SUBAPPLICATION logiBUS_QXA_OPC (* logiBUS DQ Kanal: OPC-UA Read/Write (generisch, ein Kanal, ohne VT-Button/Hintergrundfarbe - fuer Module ohne ISOBUS/VT-Anbindung) *)
  (* Standard: 61499-2 *)
  (* Version 1.0, 2026-08-27, franz, Meisterschulen am Ostbahnhof *)
  PACKAGE MyLib::sys;
  IMPORT logiBUS::io::DQ::logiBUS_DO;
  IMPORT logiBUS::io::DQ::logiBUS_DO_S;
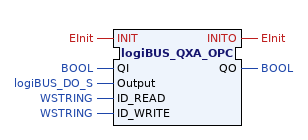
  EVENT_INPUT
    INIT : EInit; (* Initialization Request *)
  END_EVENT
  EVENT_OUTPUT
    INITO : EInit; (* Initialization Confirm *)
  END_EVENT
  VAR_INPUT
    QI : BOOL := TRUE; (* Quality Input - TRUE to enable service *)
    Output : logiBUS::io::DQ::logiBUS_DO_S := logiBUS_DO::Invalid; (* Identify the Output Output_Q1..Q12 *)
    ID_READ : WSTRING; (* OPC-UA Subscribe-Key (schreibbar) *)
    ID_WRITE : WSTRING; (* OPC-UA Publish-Key (lesbar) *)
  END_VAR
  VAR_OUTPUT
    QO : BOOL; (* Quality Output - TRUE if service executed successfully *)
  END_VAR
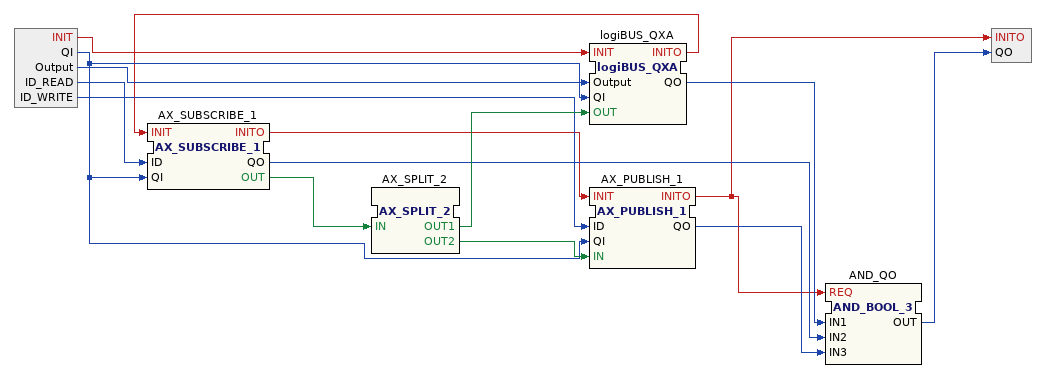
  FBS
    logiBUS_QXA : logiBUS::io::DQ::logiBUS_QXA;
    AX_SUBSCRIBE_1 : adapter::net::AX_SUBSCRIBE_1;
    AX_SPLIT_2 : adapter::events::unidirectional::AX_SPLIT_2;
    AX_PUBLISH_1 : adapter::net::AX_PUBLISH_1;
    AND_QO : iec61131::booleanOperators::AND_BOOL_3;
  END_FBS
  EVENT_CONNECTIONS
    INIT TO logiBUS_QXA.INIT;
    logiBUS_QXA.INITO TO AX_SUBSCRIBE_1.INIT;
    AX_SUBSCRIBE_1.INITO TO AX_PUBLISH_1.INIT;
    AX_PUBLISH_1.INITO TO INITO;
    AX_PUBLISH_1.INITO TO AND_QO.REQ;
  END_CONNECTIONS
  DATA_CONNECTIONS
    Output TO logiBUS_QXA.Output;
    ID_READ TO AX_SUBSCRIBE_1.ID;
    ID_WRITE TO AX_PUBLISH_1.ID;
    QI TO logiBUS_QXA.QI;
    QI TO AX_SUBSCRIBE_1.QI;
    QI TO AX_PUBLISH_1.QI;
    logiBUS_QXA.QO TO AND_QO.IN1;
    AX_SUBSCRIBE_1.QO TO AND_QO.IN2;
    AX_PUBLISH_1.QO TO AND_QO.IN3;
    AND_QO.OUT TO QO;
  END_CONNECTIONS
  ADAPTER_CONNECTIONS
    AX_SUBSCRIBE_1.OUT TO AX_SPLIT_2.IN;
    AX_SPLIT_2.OUT1 TO logiBUS_QXA.OUT;
    AX_SPLIT_2.OUT2 TO AX_PUBLISH_1.IN;
  END_CONNECTIONS
END_SUBAPPLICATION
